(* IEC 61131-3 sources: plc-st-coding-agent/progress/evidence/f14_v2_public_20261112b/jobs/custom_deepseek-v4pro, 6 files *)

(* ---- public-easy-01.candidate_01.st ---- *)
FUNCTION_BLOCK FillingLineControl
VAR_INPUT
    bottleSensor : BOOL;
    cleaningConfirmButton : BOOL;
    fillingConfirmButton : BOOL;
    cappingConfirmButton : BOOL;
    packingConfirmButton : BOOL;
    finishedButton : BOOL;
END_VAR

VAR_OUTPUT
    Pump_Motor : BOOL;
    Filling_Valve : BOOL;
    Capping_Machine : BOOL;
    Packing_Machine : BOOL;
    Completion_Light : BOOL;
END_VAR

VAR
    stepState : INT := 0;
    lastCleaningConfirmButton : BOOL := FALSE;
    lastFillingConfirmButton : BOOL := FALSE;
    lastCappingConfirmButton : BOOL := FALSE;
    lastPackingConfirmButton : BOOL := FALSE;
    lastFinishedButton : BOOL := FALSE;
    cleaningConfirmR : BOOL;
    fillingConfirmR : BOOL;
    cappingConfirmR : BOOL;
    packingConfirmR : BOOL;
    finishedR : BOOL;
END_VAR

cleaningConfirmR := cleaningConfirmButton AND NOT lastCleaningConfirmButton;
fillingConfirmR := fillingConfirmButton AND NOT lastFillingConfirmButton;
cappingConfirmR := cappingConfirmButton AND NOT lastCappingConfirmButton;
packingConfirmR := packingConfirmButton AND NOT lastPackingConfirmButton;
finishedR := finishedButton AND NOT lastFinishedButton;

CASE stepState OF
    0:
        IF bottleSensor THEN
            stepState := 1;
        END_IF;
    1:
        IF cleaningConfirmR THEN
            stepState := 2;
        END_IF;
    2:
        IF fillingConfirmR THEN
            stepState := 3;
        END_IF;
    3:
        IF cappingConfirmR THEN
            stepState := 4;
        END_IF;
    4:
        IF packingConfirmR THEN
            stepState := 5;
        END_IF;
    5:
        IF finishedR THEN
            stepState := 0;
        END_IF;
END_CASE;

Pump_Motor := (stepState = 1);
Filling_Valve := (stepState = 2);
Capping_Machine := (stepState = 3);
Packing_Machine := (stepState = 4);
Completion_Light := (stepState = 5);

lastCleaningConfirmButton := cleaningConfirmButton;
lastFillingConfirmButton := fillingConfirmButton;
lastCappingConfirmButton := cappingConfirmButton;
lastPackingConfirmButton := packingConfirmButton;
lastFinishedButton := finishedButton;

END_FUNCTION_BLOCK

(* ---- public-easy-01.candidate_02.st ---- *)
FUNCTION_BLOCK FillingLineControl
VAR_INPUT
    bottleSensor : BOOL;
    cleaningConfirmButton : BOOL;
    fillingConfirmButton : BOOL;
    cappingConfirmButton : BOOL;
    packingConfirmButton : BOOL;
    finishedButton : BOOL;
END_VAR

VAR_OUTPUT
    Pump_Motor : BOOL;
    Filling_Valve : BOOL;
    Capping_Machine : BOOL;
    Packing_Machine : BOOL;
    Completion_Light : BOOL;
END_VAR

VAR
    stepState : INT := 0;

    lastBottleSensor : BOOL := FALSE;
    lastCleaningConfirmButton : BOOL := FALSE;
    lastFillingConfirmButton : BOOL := FALSE;
    lastCappingConfirmButton : BOOL := FALSE;
    lastPackingConfirmButton : BOOL := FALSE;
    lastFinishedButton : BOOL := FALSE;

    bottleSensorR : BOOL;
    cleaningConfirmR : BOOL;
    fillingConfirmR : BOOL;
    cappingConfirmR : BOOL;
    packingConfirmR : BOOL;
    finishedR : BOOL;
END_VAR

(* 上升沿检测 *)
bottleSensorR := bottleSensor AND NOT lastBottleSensor;
cleaningConfirmR := cleaningConfirmButton AND NOT lastCleaningConfirmButton;
fillingConfirmR := fillingConfirmButton AND NOT lastFillingConfirmButton;
cappingConfirmR := cappingConfirmButton AND NOT lastCappingConfirmButton;
packingConfirmR := packingConfirmButton AND NOT lastPackingConfirmButton;
finishedR := finishedButton AND NOT lastFinishedButton;

(* 步骤状态机 *)
CASE stepState OF
    0: (* 等待瓶子到达 *)
        IF bottleSensorR THEN
            stepState := 1;
        END_IF;

    1: (* 清洁 *)
        IF cleaningConfirmR THEN
            stepState := 2;
        END_IF;

    2: (* 填充 *)
        IF fillingConfirmR THEN
            stepState := 3;
        END_IF;

    3: (* 封盖 *)
        IF cappingConfirmR THEN
            stepState := 4;
        END_IF;

    4: (* 包装 *)
        IF packingConfirmR THEN
            stepState := 5;
        END_IF;

    5: (* 完成指示 *)
        IF finishedR THEN
            stepState := 0;
        END_IF;
END_CASE;

(* 输出分配 *)
Pump_Motor := (stepState = 1);
Filling_Valve := (stepState = 2);
Capping_Machine := (stepState = 3);
Packing_Machine := (stepState = 4);
Completion_Light := (stepState = 5);

(* 更新上一次输入状态 *)
lastBottleSensor := bottleSensor;
lastCleaningConfirmButton := cleaningConfirmButton;
lastFillingConfirmButton := fillingConfirmButton;
lastCappingConfirmButton := cappingConfirmButton;
lastPackingConfirmButton := packingConfirmButton;
lastFinishedButton := finishedButton;

END_FUNCTION_BLOCK

(* ---- public-easy-02.candidate_01.st ---- *)
FUNCTION_BLOCK FB
VAR_INPUT
    value : DWORD;
END_VAR
VAR_OUTPUT
    hasChanged : BOOL;
    hasRisingEdges : BOOL;
    risingBits : DWORD;
    noOfRisingBits : USINT;
    hasFallingEdges : BOOL;
    fallingBits : DWORD;
    noOfFallingBits : USINT;
END_VAR
VAR
    lastValue : DWORD;
    firstRun : BOOL := TRUE;
    i : INT;
    mask : DWORD;
    countRise : USINT;
    countFall : USINT;
END_VAR

IF firstRun THEN
    lastValue := value;
    firstRun := FALSE;
    hasChanged := FALSE;
    hasRisingEdges := FALSE;
    risingBits := 0;
    noOfRisingBits := 0;
    hasFallingEdges := FALSE;
    fallingBits := 0;
    noOfFallingBits := 0;
    RETURN;
END_IF;

hasChanged := (value <> lastValue);
risingBits := (NOT lastValue) AND value;
fallingBits := lastValue AND (NOT value);
hasRisingEdges := (risingBits <> 0);
hasFallingEdges := (fallingBits <> 0);

countRise := 0;
FOR i := 0 TO 31 DO
    mask := SHL(DWORD#1, i);
    IF (risingBits AND mask) <> 0 THEN
        countRise := countRise + 1;
    END_IF;
END_FOR;
noOfRisingBits := countRise;

countFall := 0;
FOR i := 0 TO 31 DO
    mask := SHL(DWORD#1, i);
    IF (fallingBits AND mask) <> 0 THEN
        countFall := countFall + 1;
    END_IF;
END_FOR;
noOfFallingBits := countFall;

lastValue := value;

END_FUNCTION_BLOCK

(* ---- public-easy-02.candidate_02.st ---- *)
FUNCTION_BLOCK FB
VAR_INPUT
    value : DWORD;
END_VAR
VAR_OUTPUT
    hasChanged : BOOL;
    hasRisingEdges : BOOL;
    risingBits : DWORD;
    noOfRisingBits : USINT;
    hasFallingEdges : BOOL;
    fallingBits : DWORD;
    noOfFallingBits : USINT;
END_VAR
VAR
    lastValue : DWORD := 0;
    i : INT;
    countRise : USINT;
    countFall : USINT;
END_VAR

risingBits := (NOT lastValue) AND value;
fallingBits := lastValue AND (NOT value);
hasChanged := (value <> lastValue);
hasRisingEdges := (risingBits <> 0);
hasFallingEdges := (fallingBits <> 0);

countRise := 0;
FOR i := 0 TO 31 DO
    IF (risingBits AND SHL(DWORD#1, i)) <> 0 THEN
        countRise := countRise + 1;
    END_IF;
END_FOR;
noOfRisingBits := countRise;

countFall := 0;
FOR i := 0 TO 31 DO
    IF (fallingBits AND SHL(DWORD#1, i)) <> 0 THEN
        countFall := countFall + 1;
    END_IF;
END_FOR;
noOfFallingBits := countFall;

lastValue := value;

END_FUNCTION_BLOCK

(* ---- public-easy-03.candidate_01.st ---- *)
FUNCTION_BLOCK AlarmHandler
VAR_INPUT
    Value : REAL;
    hiLevel : REAL;
    loLevel : REAL;
    hystWindow : REAL;
END_VAR
VAR_OUTPUT
    hiAlarm : BOOL;
    loAlarm : BOOL;
    error : BOOL;
    status : WORD;
END_VAR
VAR
END_VAR

BEGIN
    error := FALSE;
    status := 0;

    IF loLevel >= hiLevel THEN
        error := TRUE;
        status := 16#8001;
        RETURN;
    ELSIF hystWindow >= (hiLevel - loLevel) THEN
        error := TRUE;
        status := 16#8002;
        RETURN;
    END_IF;

    // High limit alarm with hysteresis
    IF Value > hiLevel THEN
        hiAlarm := TRUE;
    ELSIF Value < (hiLevel - hystWindow) THEN
        hiAlarm := FALSE;
    END_IF;

    // Low limit alarm with hysteresis
    IF Value < loLevel THEN
        loAlarm := TRUE;
    ELSIF Value > (loLevel + hystWindow) THEN
        loAlarm := FALSE;
    END_IF;
END_FUNCTION_BLOCK

(* ---- public-easy-03.candidate_02.st ---- *)
FUNCTION_BLOCK AlarmHandler
VAR_INPUT
    Value : REAL;
    hiLevel : REAL;
    loLevel : REAL;
    hystWindow : REAL;
END_VAR
VAR_OUTPUT
    hiAlarm : BOOL;
    loAlarm : BOOL;
    error : BOOL;
    status : WORD;
END_VAR
VAR
END_VAR

BEGIN
    THIS^.error := FALSE;
    THIS^.status := 0;

    IF loLevel >= hiLevel THEN
        THIS^.error := TRUE;
        THIS^.status := 16#8001;
        RETURN;
    ELSIF hystWindow >= (hiLevel - loLevel) THEN
        THIS^.error := TRUE;
        THIS^.status := 16#8002;
        RETURN;
    END_IF;

    // High limit alarm with hysteresis
    IF Value > hiLevel THEN
        hiAlarm := TRUE;
    ELSIF Value < (hiLevel - hystWindow) THEN
        hiAlarm := FALSE;
    END_IF;

    // Low limit alarm with hysteresis
    IF Value < loLevel THEN
        loAlarm := TRUE;
    ELSIF Value > (loLevel + hystWindow) THEN
        loAlarm := FALSE;
    END_IF;
END_FUNCTION_BLOCK
